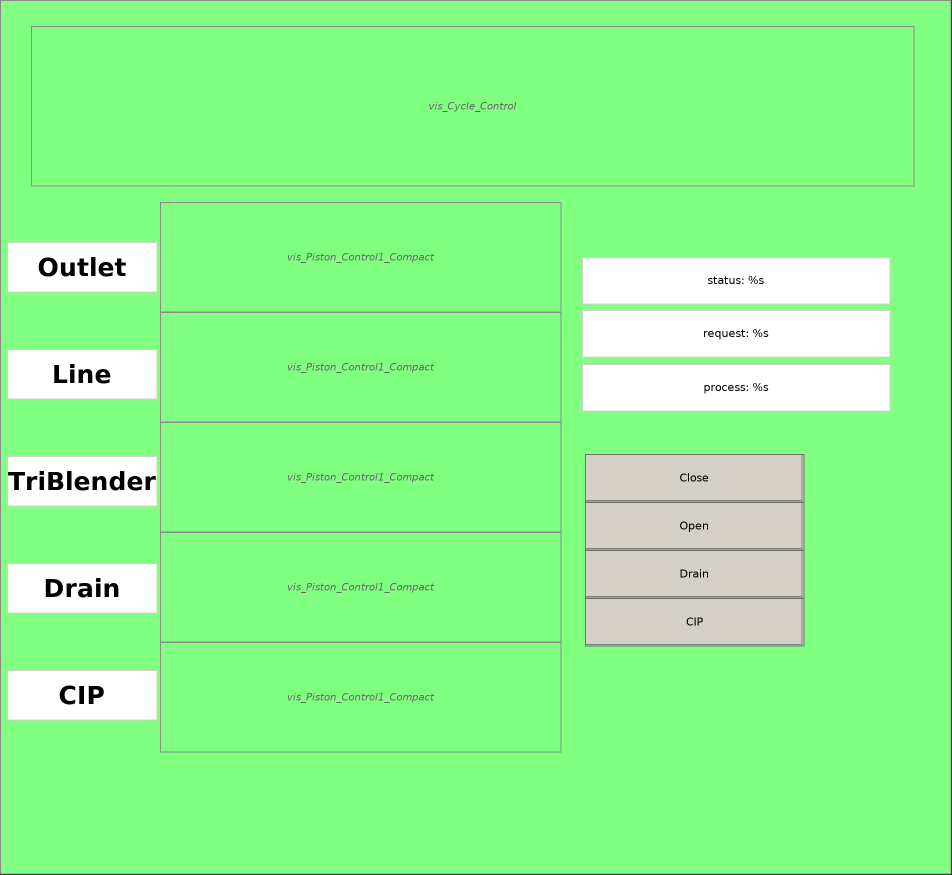
VISUALIZATION vis_FB_Tank_Target  // 952x875
VAR_IN_OUT
	fb: FB_Tank_Target;
END_VAR
    Rectangle (0,0 952x875)
    Frame (160,202 401x110)
        shows vis_Piston_Control1_Compact(stPis := fb.stPis_Outlet)
    Frame (160,312 401x110)
        shows vis_Piston_Control1_Compact(stPis := fb.stPis_Line)
    Frame (160,422 401x110)
        shows vis_Piston_Control1_Compact(stPis := fb.stPis_TriBlender)
    Frame (160,532 401x110)
        shows vis_Piston_Control1_Compact(stPis := fb.stPis_Drain)
    Frame (160,642 401x110)
        shows vis_Piston_Control1_Compact(stPis := fb.stPis_CIP)
    Frame (31,26 883x160)
        shows vis_Cycle_Control(fb := fb, sName := 'Tank Target Interface')
    Textfield (582,257 308x47), "status: %s", text variable: fb.eStatus
    Button (585,454 219x48), "Close"
        OnMouseClick: execute { fb.eReq:=E_Tank_Target.eClose; }
    Textfield (582,310 308x47), "request: %s", text variable: fb.eReq
    Textfield (582,364 308x47), "process: %s", text variable: fb.eProcess
    Button (585,502 219x48), "Open"
        OnMouseClick: execute { fb.eReq:=E_Tank_Target.eOpen; }
    Button (585,550 219x48), "Drain"
        OnMouseClick: execute { fb.eReq:=E_Tank_Target.eDrain; }
    Button (585,598 219x48), "CIP"
        OnMouseClick: execute { fb.eReq:=E_Tank_Target.eCIP; }
    Textfield (7,242 150x50), "Outlet"
    Textfield (7,349 150x50), "Line"
    Textfield (7,456 150x50), "TriBlender"
    Textfield (7,563 150x50), "Drain"
    Textfield (7,670 150x50), "CIP"
END_VISUALIZATION

(* stored: Version 1.1.0.1, ProductVersion 3.1.4024.12
   Visu vis_FB_Tank_Target: Id {53cba01e-dc91-4db1-a16f-5213b07acfcb} *)
